(* IEC 61131-3 sources: kns-pump-station/src/POUs/Field/FB_VfdAdapter_Cond, 5 files *)

(* ---- FB_VfdAdapter_Cond.decl.st ---- *)
// Назначение: адаптер ПЧ по условной карте регистров (не карта реального производителя, ARCHITECTURE,
//             раздел 12): Decode разбирает слово состояния STW и фактическую частоту FACT для PL.FB_MotorVfd,
//             Encode собирает слово управления CTW (бит сброса аварии, пока xQReset) и задание частоты FREF.
//             Пуск — проводом (P10n_RUN), бит пуска в CTW не используется. Без связи слово состояния
//             недостоверно: готовность, работа, авария, предупреждение, местное — FALSE, скорость — последняя
//             принятая; частоту ПЧ задаёт его сторожевой таймер (04 §12). Другая модель ПЧ — другой адаптер
//             с теми же выходами.
// Автор:      kr0nsch
// Версия:     0.1.0
// Документ:   docs/DESIGN.md, раздел 8.2; docs/ARCHITECTURE.md, раздел 12
FUNCTION_BLOCK FB_VfdAdapter_Cond
VAR_OUTPUT
    xCommOk       : BOOL;           // xSlaveOk последнего Decode
    xReady        : BOOL;           // STW.0 (при связи; без связи — FALSE)
    xRunning      : BOOL;           // STW.1
    xFault        : BOOL;           // STW.2
    xWarning      : BOOL;           // STW.3 (HMI)
    xRemote       : BOOL;           // STW.4 (HMI)
    rSpeedAct_pct : REAL;           // FACT / VFD_COUNTS_PER_PCT; без связи — последнее значение
    wCtw          : WORD;           // слово управления (Encode)
    uiFref        : UINT;           // задание частоты, 0,01 Гц (Encode)
END_VAR

(* ---- Decode.method.decl.st ---- *)
// Разобрать регистры чтения ПЧ (FC3 100, 101) и состояние обмена со слейвом
METHOD Decode
VAR_INPUT
    wStw     : WORD;                // слово состояния (GVL_IO.wP10n_STW)
    uiFact   : UINT;                // фактическая частота, 0,01 Гц (GVL_IO.uiP10n_FACT)
    xSlaveOk : BOOL;                // обмен со слейвом исправен (GVL_IO.xMbOk_RS485_1_Sn)
END_VAR

(* ---- Decode.method.impl.st ---- *)
xCommOk := xSlaveOk;
IF xSlaveOk THEN
    xReady := (wStw AND GVL_Const.VFD_STW_READY) <> 0;
    xRunning := (wStw AND GVL_Const.VFD_STW_RUNNING) <> 0;
    xFault := (wStw AND GVL_Const.VFD_STW_FAULT) <> 0;
    xWarning := (wStw AND GVL_Const.VFD_STW_WARNING) <> 0;
    xRemote := (wStw AND GVL_Const.VFD_STW_REMOTE) <> 0;
    rSpeedAct_pct := UINT_TO_REAL(uiFact) / GVL_Const.VFD_COUNTS_PER_PCT;
ELSE
    // регистры без связи замирают: слово состояния недостоверно, скорость — последняя принятая
    xReady := FALSE;
    xRunning := FALSE;
    xFault := FALSE;
    xWarning := FALSE;
    xRemote := FALSE;
END_IF

(* ---- Encode.method.decl.st ---- *)
// Собрать регистры записи ПЧ (FC16 0, 1): бит сброса аварии, пока xQReset (импульс библиотеки 1 с длиннее
// цикла записи Modbus), задание частоты — LIMIT(0, rSpeedRef_pct, 100) · VFD_COUNTS_PER_PCT с округлением;
// неконечное задание — 0
METHOD Encode
VAR_INPUT
    xQReset       : BOOL;           // импульс сброса аварии ПЧ (GVL_IO.xP10n_VfdQReset ← fbP10n.xQReset)
    rSpeedRef_pct : REAL;           // задание на ПЧ, % (GVL_IO.rP10n_SpeedRef_pct ← fbP10n.rSpeedRef_pct)
END_VAR

(* ---- Encode.method.impl.st ---- *)
wCtw := SEL(xQReset, 0, GVL_Const.VFD_CTW_RESET);
IF PL.F_IsFinite(rIn := rSpeedRef_pct) THEN
    uiFref := REAL_TO_UINT(LIMIT(0.0, rSpeedRef_pct, PL.GVL_Const.PCT_FULL) * GVL_Const.VFD_COUNTS_PER_PCT);
ELSE
    uiFref := 0;
END_IF
